(* IEC 61131-3 sources: nautilus/examples/alarms, 3 files *)

(* ---- blocks.st ---- *)
(* A root .st file with no PROGRAM is a library: it is in scope for every
   task's compile, so `type: AnalogInput` in the manifest resolves against
   it — and so an alarm rule can say `match: {type: AnalogInput, member:
   HH}` and mean this. *)

TYPE
  AnalogInput : STRUCT
    PV : REAL;   (* the measurement *)
    HH : BOOL;   (* the four limit bits the alarm rules claim *)
    H  : BOOL;
    L  : BOOL;
    LL : BOOL;
  END_STRUCT;
END_TYPE

(* ---- program.st ---- *)
PROGRAM Annunciate
(* The bits, computed in control logic at scan rate. That is the whole
   division of labour: comparing a measurement to a limit is control, and
   deciding whether a person has to be told about it — and whether they
   have seen it yet — is alarm management, which lives in the host's alarm
   engine, not here. Nothing in this program knows an alarm engine exists. *)
VAR_EXTERNAL
    RTU9_WEL15_FIT_001 : AnalogInput;
    RTU9_TNK01_LIT_001 : AnalogInput;

    FlowHH  : REAL;  FlowH  : REAL;  FlowL  : REAL;  FlowLL  : REAL;
    LevelHH : REAL;  LevelH : REAL;  LevelL : REAL;  LevelLL : REAL;

    RTU9__Online : BOOL;
    RTU9_AnyAlm  : BOOL;
END_VAR

RTU9_WEL15_FIT_001.HH := RTU9_WEL15_FIT_001.PV > FlowHH;
RTU9_WEL15_FIT_001.H  := RTU9_WEL15_FIT_001.PV > FlowH;
RTU9_WEL15_FIT_001.L  := RTU9_WEL15_FIT_001.PV < FlowL;
RTU9_WEL15_FIT_001.LL := RTU9_WEL15_FIT_001.PV < FlowLL;

RTU9_TNK01_LIT_001.HH := RTU9_TNK01_LIT_001.PV > LevelHH;
RTU9_TNK01_LIT_001.H  := RTU9_TNK01_LIT_001.PV > LevelH;
RTU9_TNK01_LIT_001.L  := RTU9_TNK01_LIT_001.PV < LevelL;
RTU9_TNK01_LIT_001.LL := RTU9_TNK01_LIT_001.PV < LevelLL;

(* The site rollup an overview screen shows. It is gated on the node being
   online for the same reason every alarm definition is: a dead edge node
   holds its last values, so an ungated rollup would stay lit forever. *)
RTU9_AnyAlm := RTU9__Online AND (
      RTU9_WEL15_FIT_001.HH OR RTU9_WEL15_FIT_001.L
   OR RTU9_TNK01_LIT_001.HH OR RTU9_TNK01_LIT_001.L);

END_PROGRAM

(* ---- sim.st ---- *)
PROGRAM Sim
(* The plant, so `nautilus run` shows alarms coming and going without any
   field hardware. Acceptance tests suspend this task and drive the
   measurements themselves — freezing the thing that would otherwise fight
   the test is what turns a closed loop into an open-loop assertion. *)
VAR_EXTERNAL
    RTU9_WEL15_FIT_001 : AnalogInput;
    RTU9_TNK01_LIT_001 : AnalogInput;
    RTU9_WEL15_INT_001_YA : BOOL;
    SimDtS : REAL;
END_VAR
VAR
    t : REAL := 0.0;
END_VAR

t := t + SimDtS;
IF t > 120.0 THEN t := 0.0; END_IF;

RTU9_WEL15_FIT_001.PV := t;           (* ramps up through the flow HH limit *)
RTU9_TNK01_LIT_001.PV := 120.0 - t;   (* and the tank drains through its L  *)
RTU9_WEL15_INT_001_YA := t > 110.0;   (* a standalone contact, briefly made  *)

END_PROGRAM
